TYPE ST_AlarmRef_1 :
STRUCT
	stControl				:ST_AlarmOut;
	stManual				:ST_AlarmOut;
	//stMaintenance			:ST_AlarmOut;
	stHome					:ST_AlarmOut;
	stAuto					:ST_AlarmOut;
END_STRUCT
END_TYPE

(* stored: Version 1.1.0.1, ProductVersion 3.1.4024.15
   DUT ST_AlarmRef_1: Id {1e23baa9-8b90-45a9-a3fe-ef9bd12e25c4} *)
